Staubli VAL3: MoveCirc.pgx

program MoveCirc(num x_nX, num x_nY, num x_nZ, num x_nRx, num x_nRy, num x_nRz, num x_nX2, num x_nY2, num x_nZ2, num x_nRx2, num x_nRy2, num x_nRz2)
begin
  pPointRx.trsf.x = x_nX
  pPointRx.trsf.y = x_nY
  pPointRx.trsf.z = x_nZ
  pPointRx.trsf.rx = x_nRx
  pPointRx.trsf.ry = x_nRy
  pPointRx.trsf.rz = x_nRz
  pPointRx2.trsf.x = x_nX2
  pPointRx2.trsf.y = x_nY2
  pPointRx2.trsf.z = x_nZ2
  pPointRx2.trsf.rx = x_nRx2
  pPointRx2.trsf.ry = x_nRy2
  pPointRx2.trsf.rz = x_nRz2
  movec(pPointRx,pPointRx2,tCurrentTool,mCurrentSpeed)
end
